Fanuc KAREL source: kb00071.compact.KL

PROGRAM KB00071
%STACKSIZE=65535
%PRIORITY=65535
%NOLOCKGROUP
VAR
P1 : REAL
RESULT : REAL
BEGIN
P1=1.0
RESULT=EXP(P1)
END KB00071
